// TIA Portal V20 export
// export: Created 2026-10-19T18:42:23.8027704Z, ExportSetting WithDefaults, DisplayName Totally Integrated Automation Portal, DisplayVersion V20 Update 6, DisplayName TIA Portal Openness, DisplayVersion V20 Update 6, DisplayName TIA Portal Version Control Interface, DisplayVersion V20 Update 6, DisplayName SINAMICS Startdrive Advanced, DisplayVersion V20 SP1, DisplayName SINAMICS Startdrive G130, G150, S120, S150, SINAMICS MV, G220, S200, S210, DisplayVersion V20 SP1, DisplayName SINAMICS Startdrive G110M, G120, G120C, G120D, G120P, G115D, DisplayVersion V20 SP1, DisplayName STEP 7 Professional, DisplayVersion V20 Update 6, DisplayName STEP 7 Safety, DisplayVersion V20 Update 2, DisplayName WinCC Basic/Comfort/Advanced, DisplayVersion V20 Update 6, DisplayName WinCC Unified, DisplayVersion V20 Update 6
FUNCTION_BLOCK "Stack_Lights_FB"   // FB21, SCL
{ S7_Optimized_Access := 'TRUE' }
VERSION : 0.1
// stored: AutoNumber true, IsIECCheckEnabled false, IsRetainMemResEnabled false, MemoryReserve 100, SetENOAutomatically false, UDAEnableTagReadback false
   VAR_INPUT
      System_Auto : Bool;
      Fault : Bool;
   END_VAR
   VAR_OUTPUT
      Red : Bool;
      Green : Bool;
      Orange : Bool;
   END_VAR
BEGIN
   //Commands for Stack Light

   IF #Fault THEN  // Fault = Red
       #Red := "Clock_0.5Hz";
       #Green := FALSE;
       #Orange := FALSE;
   ELSIF #System_Auto THEN  // (1)Manual = Yellow
       #Orange := FALSE;
       #Red := FALSE;
       #Green := TRUE;
   ELSIF NOT #System_Auto THEN  // (2)Semi-Auto = Blue
       #Green := FALSE;
       #Orange := TRUE;
       #Red := FALSE;
   // ELSIF #System_Auto = 3 THEN  // (3)Auto = Green
   //     #Green := FALSE;
   //     #Red := FALSE;
   //     #Yellow := TRUE;

   ELSE
       #Green := FALSE;
       #Red := FALSE;
       #Orange := FALSE;
   END_IF;
END_FUNCTION_BLOCK
